// Mitsubishi GX Works2 project: 261012_타이머실습_타이머추가응용2   PLC: Q03UDV

PROGRAM MAIN
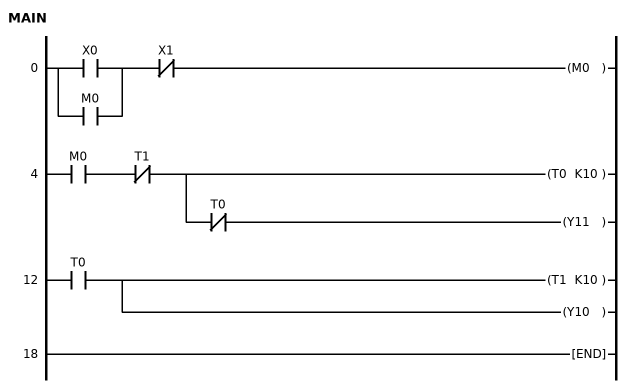
0     LD      X0
      OR      M0
      ANI     X1
      OUT     M0
4     LD      M0
      ANI     T1
      OUT     T0 K10
      ANI     T0
      OUT     Y11
12    LD      T0
      OUT     T1 K10
      OUT     Y10
18    END
END_PROGRAM
